Staubli VAL3: actionItem.dtx

public num nIOindex
public num nboolValue
public num nPulseValue
public string sIOtype
public string sValue
public bool bActive
